FUNCTION_BLOCK Name
  (* Standard: 61499-1; Description: Copyright (c) 2026 Martin Erich Jobst This program and the accompanying materials are made available under the terms of the Eclipse Public License 2.0 which is available at https://www.eclipse.org/legal/epl-2.0/ SPDX-License-Identifier: EPL-2.0 *)
  (* Version 1.0, 2026-11-18, Martin Jobst *)
  PACKAGE lib::IInterfaceElement;
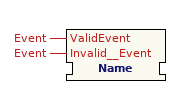
  EVENT_INPUT
    ValidEvent;
    Invalid__Event;
  END_EVENT
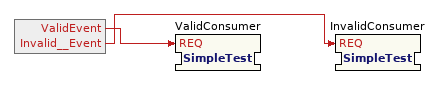
  FBS
    ValidConsumer : lib::IInterfaceElement::support::SimpleTest;
    InvalidConsumer : lib::IInterfaceElement::support::SimpleTest;
  END_FBS
  EVENT_CONNECTIONS
    ValidEvent TO ValidConsumer.REQ;
    Invalid__Event TO InvalidConsumer.REQ;
  END_CONNECTIONS
END_FUNCTION_BLOCK
